(* PLC project TBEN_L5_PLC11.project, CODESYS CODESYS V3.5 SP21 Patch 1 *)
(* stored: creationDateTime 2026-11-07T15:35:07.161101, modificationDateTime 2026-11-07T15:09:07.4034196 *)

// Định nghĩa 1 event của device (từ IODD)
TYPE ST_IolEventDef :
STRUCT
    wCode  : WORD;
    sName  : STRING(12);        // tên ngắn trên màn hình cảm biến
    wsText : WSTRING(48);       // mô tả cho HMI
    eType  : E_IolEvtType;
END_STRUCT
END_TYPE
